Staubli VAL3: ParaItem.pjx

--- ParaItem.pjx ---
Parameters version=s8.10.3Cs9_BS2093 stackSize=5000 millimeterUnit=true
Program file=start.pgx
Program file=stop.pgx
Data file=ParaItem.dtx
Type name=ifItem path=Disk://source/template/ifItem/ifItem.pjx

--- ParaItem.dtx ---
public mdesc mMdesc
public num nMoveType
public num nActionIndex
public num nPercentage
public ifItem iIfItem
  [0]
    num nSigType[3]
    num nSigIndex[3]
    num nValue[3]
    bool bANDOR[2]
public num nDelay
public num nSigValue
public bool bSafePoint

--- start.pgx ---
program start()
begin
end

--- stop.pgx ---
program stop()
begin
end
